// 书籍分拣功能块主逻辑
        // 1. 电机控制逻辑: 任何RFID检测到书籍时启动电机
        Motor := RFID1 OR RFID2 OR RFID3;

        // 2. 分拣箱控制逻辑: 根据RFID检测结果打开对应箱子，同一时间只有一个箱子打开
        // 优先级别: RFID1 > RFID2 > RFID3
        Bin1 := RFID1 AND NOT (RFID2 OR RFID3);
        Bin2 := RFID2 AND NOT (RFID1 OR RFID3);
        Bin3 := RFID3 AND NOT (RFID1 OR RFID2);

        // 形式化属性验证断言
        // 属性1: 电机状态与RFID检测结果的一致性
        ASSERT((RFID1 OR RFID2 OR RFID3) = Motor);

        // 属性2: 同一时间最多只有一个箱子打开或全部关闭
        ASSERT(
          (Bin1 AND NOT Bin2 AND NOT Bin3) OR
          (Bin2 AND NOT Bin1 AND NOT Bin3) OR
          (Bin3 AND NOT Bin1 AND NOT Bin2) OR
          (NOT Bin1 AND NOT Bin2 AND NOT Bin3)
        );

        // 属性3: 无书籍时所有设备处于关闭状态
        ASSERT(
          (RFID1 OR RFID2 OR RFID3) OR
          (NOT Motor AND NOT Bin1 AND NOT Bin2 AND NOT Bin3)
        );
